(* IEC 61131-3 sources: voltrus-explorers/crates/mt-plc-cli/tests/fixtures/ld, 2 files *)

(* ---- alarm-latch.golden.st ---- *)
PROGRAM AlarmLatch
VAR_INPUT
    X0 : BOOL;
    X1 : BOOL;
    X2 : BOOL;
    X3 : BOOL;
END_VAR
VAR_OUTPUT
    Y0 : BOOL;
END_VAR
VAR
    M0 : BOOL;
END_VAR

    IF (X0 OR X1 OR X2) THEN M0 := TRUE; END_IF;
    Y0 := M0;
    IF X3 THEN M0 := FALSE; END_IF;
END_PROGRAM

(* ---- motor-start-stop.golden.st ---- *)
PROGRAM MotorStartStop
VAR_INPUT
    X0 : BOOL;
    X1 : BOOL;
END_VAR
VAR_OUTPUT
    Y0 : BOOL;
END_VAR
VAR
    Y0 : BOOL;
END_VAR

    Y0 := (X0 AND NOT X1 OR Y0 AND NOT X1);
END_PROGRAM
